(* IEC 61131-3 sources: codesys-ai-industrial-robot-control/plc/src/Framework/FB_AlarmHandler, 5 files *)

(* ---- AcknowledgeAll.st ---- *)
// Acknowledge every alarm. Active alarms stay listed until their condition clears.
METHOD AcknowledgeAll
VAR
    eId : E_AlarmId;
END_VAR

FOR eId := E_AlarmId.EStop TO E_AlarmId.QueueOverflow DO
    aAlarms[eId].xAcked := TRUE;
END_FOR

(* ---- Clear.st ---- *)
METHOD Clear
VAR_INPUT
    eId : E_AlarmId;
END_VAR

aAlarms[eId].xActive := FALSE;

(* ---- GetAlarm.st ---- *)
METHOD GetAlarm : ST_Alarm
VAR_INPUT
    eId : E_AlarmId;
END_VAR

GetAlarm := aAlarms[eId];

(* ---- Raise.st ---- *)
METHOD Raise
VAR_INPUT
    eId : E_AlarmId;
END_VAR

IF eId = E_AlarmId.None OR aAlarms[eId].xActive THEN
    RETURN;
END_IF
aAlarms[eId].eClass := GVL_AlarmDefs.aDefs[eId].eClass;
aAlarms[eId].xActive := TRUE;
aAlarms[eId].xAcked := FALSE;
aAlarms[eId].tRaised := TIME();
eNewest := eId;

(* ---- RaiseEvent.st ---- *)
METHOD RaiseEvent
VAR_INPUT
    eId : E_AlarmId;
END_VAR

IF eId = E_AlarmId.None THEN
    RETURN;
END_IF
aAlarms[eId].eClass := GVL_AlarmDefs.aDefs[eId].eClass;
aAlarms[eId].xActive := FALSE;
aAlarms[eId].xAcked := FALSE;
aAlarms[eId].tRaised := TIME();
eNewest := eId;
